(* IEC 61131-3 sources: kns-pump-station/tests/POUs/Model/FB_InflowProfile_Test, 8 files *)

(* ---- FB_InflowProfile_Test.decl.st ---- *)
// Назначение: набор coUnit для FB_InflowProfile — суточный профиль притока: значения в точках и между
//             ними, переход через полночь, среднее за сутки, неконечные входы. Ожидаемые значения — эталон
//             tools_project/plant_reference.py, сценарий inflow.profile (профиль ST_SimCfg по умолчанию).
// Автор:      kr0nsch
// Версия:     0.1.0
// Документ:   docs/DESIGN.md, разделы 11.3, 14.1
FUNCTION_BLOCK FB_InflowProfile_Test EXTENDS coUnit.FB_TestSuite
VAR CONSTANT
    R_AVG_M3H : REAL := 70.0;         // stSimCfg.rInflowAvg_m3h по умолчанию
    R_EPS : REAL := 1.0E-4;           // допуск REAL для значений порядка 100
    UI_SAMPLES : UINT := 96;          // отсчётов за сутки (через 15 мин)
    R_SAMPLE_H : REAL := 0.25;
    DW_NAN : DWORD := 16#7FC00000;
END_VAR

(* ---- DefaultsMatchProfilePoints.method.decl.st ---- *)
// Профиль по умолчанию: в точке 8 ч — 1,60 · 70 = 112 м³/ч, в 3 ч — 0,38 · 70 = 26,6 м³/ч (06 §5.4: 27…112).
METHOD PRIVATE DefaultsMatchProfilePoints
VAR
    fbDut : FB_InflowProfile;   // проверяемый ФБ
    stCfg : ST_SimCfg;          // профиль по умолчанию
END_VAR

(* ---- InterpolatesBetweenHours.method.decl.st ---- *)
// Между точками — линейно: 8:30 — (1,60 + 1,50)/2 · 70 = 108,5 м³/ч; 8:45 — 1,525.
METHOD PRIVATE InterpolatesBetweenHours
VAR
    fbDut : FB_InflowProfile;   // проверяемый ФБ
    stCfg : ST_SimCfg;          // профиль по умолчанию
END_VAR

(* ---- MeanIsAverage.method.decl.st ---- *)
// Среднее за сутки (96 отсчётов через 15 мин) равно rAverage_m3h: среднее точек профиля — 1,0.
METHOD PRIVATE MeanIsAverage
VAR
    fbDut : FB_InflowProfile;   // проверяемый ФБ
    stCfg : ST_SimCfg;          // профиль по умолчанию
    uiI : UINT;
    rSum : REAL;               // сумма притока по отсчётам
END_VAR

(* ---- MeanIsAverage.method.impl.st ---- *)
coUnit.TEST('InflowProfile_MeanIsAverage');

FOR uiI := 0 TO UI_SAMPLES - 1 DO
    fbDut(rTimeOfDay_h := UINT_TO_REAL(uiI) * R_SAMPLE_H, rAverage_m3h := R_AVG_M3H, arProfile := stCfg.arDailyProfile);
    rSum := rSum + fbDut.rInflow_m3h;
END_FOR
// ref: inflow.profile.mean_factor (= 1,0)
AssertEquals_REAL(Expected := R_AVG_M3H, Actual := rSum / UINT_TO_REAL(UI_SAMPLES), Delta := 1.0E-3,
                  Message := 'daily mean equals average inflow');

coUnit.TEST_FINISHED();

(* ---- NegativeFactorGivesZeroInflow.method.decl.st ---- *)
// Отрицательный множитель (ошибка ввода профиля) не даёт отрицательного притока.
METHOD PRIVATE NegativeFactorGivesZeroInflow
VAR
    fbDut : FB_InflowProfile;   // проверяемый ФБ
    stCfg : ST_SimCfg;          // профиль по умолчанию
END_VAR

(* ---- NonFiniteInputsSafe.method.decl.st ---- *)
// Неконечное время суток — как 0 ч; неконечный средний приток — приток 0; выходы конечны.
METHOD PRIVATE NonFiniteInputsSafe
VAR
    fbDut : FB_InflowProfile;   // проверяемый ФБ
    stCfg : ST_SimCfg;          // профиль по умолчанию
    uBits : PL.U_RealBits;
END_VAR

(* ---- WrapsAtMidnight.method.decl.st ---- *)
// После 23 ч — к точке 0: 23:30 — (0,70 + 0,55)/2 = 0,625; время вне суток приводится по модулю:
// 24,25 ч = 0,25 ч; −0,5 ч = 23,5 ч.
METHOD PRIVATE WrapsAtMidnight
VAR
    fbDut : FB_InflowProfile;   // проверяемый ФБ
    stCfg : ST_SimCfg;          // профиль по умолчанию
    rRef : REAL;               // множитель в 0:15
END_VAR
